Fanuc KAREL source: KT00347.KL

PROGRAM KT00347
%NOLOCKGROUP
VAR
  P1: POSITION
  P2: POSITION
  OUT: BOOLEAN
BEGIN
  OUT = P1 < P2
END KT00347
